// The command inputs bStop/bPark/bPower/bReset of FB_TelescopeControl (IAG50cm) are edge-triggered like the methods and are never
// written by the block; the block works on the request latches bStopActive/bParkActive/bPowerActive/bResetActive.
// Plan: BROTLib specs/plans/2026-11-09-iag50cm-command-model-unification.md, steps 1a/1b. One rig per test, one Scan() per PLC cycle.
FUNCTION_BLOCK IagCommandInputs_Tests EXTENDS TcUnit.FB_TestSuite
VAR
END_VAR

Held_Stop_Input_Stops_Once();
Park_Input_Edge_Parks_Like_Park();
Stop_Method_And_Input_Edge_In_One_Scan_Count_Once();
Power_Input_Is_Not_Written_By_The_Block();
Held_Slew_Input_Starts_The_Slew_Once();
Slew_Input_Falling_Does_Not_Abort_The_Slew();
Slew_Method_And_Input_Edge_In_One_Scan_Count_Once();
Slew_Input_In_The_Scan_Of_A_New_Error_Is_Rejected();
Track_Method_And_Track_Input_In_One_Scan_Count_Once();

// A held stop input is one command: one stop transaction, never repeated, never cleared by the block (IAG50cm command model step 1a).
METHOD PRIVATE Held_Stop_Input_Stops_Once
VAR_INST
	rig			: FB_IagRig;
	nStep		: INT;
	nCycles		: UINT;
	nEdges		: UINT;
	sTest		: STRING(80);
END_VAR
TEST('Held_Stop_Input_Stops_Once');
sTest := 'Held_Stop_Input_Stops_Once: ';
IF nStep >= 90 THEN
	RETURN;
END_IF
rig.Scan();
nCycles := nCycles + 1;
CASE nStep OF
0:	// wait for the clock, then power on
	IF rig.ClockValid THEN
		rig.fbTel.Init();
		nStep := 10;
		nCycles := 0;
	ELSIF nCycles > 2000 THEN
		AssertTrue(Condition := FALSE, Message := 'the astronomical clock never became valid');
		F_Note(bFailed := TRUE, sText := CONCAT(sTest, 'the astronomical clock never became valid'));
		nStep := 99;
		TEST_FINISHED();
	END_IF
10:	// wait until the startup has finished (READY_STATE 1.0)
	IF rig.Online THEN
		rig.fbTel.Slew(fAzimuth := 180.0, fAltitude := 45.0);
		nStep := 20;
		nCycles := 0;
	ELSIF nCycles > 1500 THEN
		AssertTrue(Condition := FALSE, Message := 'the mock telescope did not reach READY_STATE 1.0');
		F_Note(bFailed := TRUE, sText := CONCAT(sTest, 'the mock telescope did not reach READY_STATE 1.0'));
		nStep := 99;
		TEST_FINISHED();
	END_IF
20:	// an axis is moving
	IF rig.fbHa.MoveAxis OR rig.fbDec.MoveAxis THEN
		nCycles := 0;
		nStep := 30;
	ELSIF nCycles > 300 THEN
		AssertTrue(Condition := FALSE, Message := 'the slew did not start an axis move');
		F_Note(bFailed := TRUE, sText := CONCAT(sTest, 'the slew did not start an axis move'));
		nStep := 99;
		TEST_FINISHED();
	END_IF
30:	// a few scans of motion, then hold the stop INPUT (an ADS write, not the method)
	IF nCycles >= 5 THEN
		rig.SetStopInput(TRUE);
		nStep := 40;
		nCycles := 0;
	END_IF
40:	// the stop has settled: note the stop edges, keep holding the input
	IF NOT rig.fbTel.bStopActive AND rig.fbTel.bStopped AND nCycles > 5 THEN
		nEdges := rig.fbHa.nStopEdges + rig.fbDec.nStopEdges;
		AssertTrue(Condition := nEdges = 1, Message := 'the held input sent one stop to the moving axis');
		F_Note(bFailed := NOT (nEdges = 1), sText := CONCAT(sTest, 'the held input sent one stop to the moving axis'));
		nStep := 50;
		nCycles := 0;
	ELSIF nCycles > 400 THEN
		AssertTrue(Condition := FALSE, Message := 'the stop did not settle');
		F_Note(bFailed := TRUE, sText := CONCAT(sTest, 'the stop did not settle'));
		nStep := 99;
		TEST_FINISHED();
	END_IF
50:	// 60 more scans with the input still TRUE: no second stop, the latch stays down, the input is not cleared
	IF nCycles >= 60 THEN
		AssertTrue(Condition := rig.fbHa.nStopEdges + rig.fbDec.nStopEdges = nEdges, Message := 'a held input is not a second stop');
		F_Note(bFailed := NOT (rig.fbHa.nStopEdges + rig.fbDec.nStopEdges = nEdges), sText := CONCAT(sTest, 'a held input is not a second stop'));
		AssertTrue(Condition := NOT rig.fbTel.bStopActive, Message := 'the stop latch stayed down');
		F_Note(bFailed := NOT (NOT rig.fbTel.bStopActive), sText := CONCAT(sTest, 'the stop latch stayed down'));
		AssertTrue(Condition := rig.fbTel.bStop, Message := 'the block did not clear the input');
		F_Note(bFailed := NOT (rig.fbTel.bStop), sText := CONCAT(sTest, 'the block did not clear the input'));
		AssertTrue(Condition := rig.fbFocus.nStop = 1, Message := 'one stop for the focus');
		F_Note(bFailed := NOT (rig.fbFocus.nStop = 1), sText := CONCAT(sTest, 'one stop for the focus'));
		nStep := 99;
		TEST_FINISHED();
	END_IF
END_CASE
END_METHOD

// A rising park input starts the park exactly like Park(); the finished park is not replayed from the held input.
METHOD PRIVATE Park_Input_Edge_Parks_Like_Park
VAR_INST
	rig			: FB_IagRig;
	nStep		: INT;
	nCycles		: UINT;
	nEdges		: UINT;
	sTest		: STRING(80);
END_VAR
TEST('Park_Input_Edge_Parks_Like_Park');
sTest := 'Park_Input_Edge_Parks_Like_Park: ';
IF nStep >= 90 THEN
	RETURN;
END_IF
rig.Scan();
nCycles := nCycles + 1;
CASE nStep OF
0:	// wait for the clock, then power on
	IF rig.ClockValid THEN
		rig.fbTel.Init();
		nStep := 10;
		nCycles := 0;
	ELSIF nCycles > 2000 THEN
		AssertTrue(Condition := FALSE, Message := 'the astronomical clock never became valid');
		F_Note(bFailed := TRUE, sText := CONCAT(sTest, 'the astronomical clock never became valid'));
		nStep := 99;
		TEST_FINISHED();
	END_IF
10:	// wait until the startup has finished (READY_STATE 1.0)
	IF rig.Online THEN
		rig.SetParkInput(TRUE);
		nStep := 20;
		nCycles := 0;
	ELSIF nCycles > 1500 THEN
		AssertTrue(Condition := FALSE, Message := 'the mock telescope did not reach READY_STATE 1.0');
		F_Note(bFailed := TRUE, sText := CONCAT(sTest, 'the mock telescope did not reach READY_STATE 1.0'));
		nStep := 99;
		TEST_FINISHED();
	END_IF
20:	// the edge starts the park, as Park() would
	IF rig.fbTel.bParkActive THEN
		nStep := 30;
		nCycles := 0;
	ELSIF nCycles > 10 THEN
		AssertTrue(Condition := FALSE, Message := 'the park input edge did not start the park');
		F_Note(bFailed := TRUE, sText := CONCAT(sTest, 'the park input edge did not start the park'));
		nStep := 99;
		TEST_FINISHED();
	END_IF
30:
	IF rig.fbTel.bIsParked THEN
		nStep := 40;
		nCycles := 0;
	ELSIF nCycles > 3000 THEN
		AssertTrue(Condition := FALSE, Message := 'the park did not finish');
		F_Note(bFailed := TRUE, sText := CONCAT(sTest, 'the park did not finish'));
		nStep := 99;
		TEST_FINISHED();
	END_IF
40:	// the park ended with the input still TRUE: it is not replayed and not cleared
	IF nCycles >= 30 THEN
		AssertTrue(Condition := NOT rig.fbTel.bParkActive, Message := 'the park request ended');
		F_Note(bFailed := NOT (NOT rig.fbTel.bParkActive), sText := CONCAT(sTest, 'the park request ended'));
		AssertTrue(Condition := rig.fbTel.bIsParked, Message := 'the telescope stays parked');
		F_Note(bFailed := NOT (rig.fbTel.bIsParked), sText := CONCAT(sTest, 'the telescope stays parked'));
		AssertTrue(Condition := rig.fbTel.bPark, Message := 'the block did not clear the input');
		F_Note(bFailed := NOT (rig.fbTel.bPark), sText := CONCAT(sTest, 'the block did not clear the input'));
		nStep := 99;
		TEST_FINISHED();
	END_IF
END_CASE
END_METHOD

// Stop() and a stop input edge in one scan are one command (the method sets the edge memory).
METHOD PRIVATE Stop_Method_And_Input_Edge_In_One_Scan_Count_Once
VAR_INST
	rig			: FB_IagRig;
	nStep		: INT;
	nCycles		: UINT;
	nEdges		: UINT;
	sTest		: STRING(80);
END_VAR
TEST('Stop_Method_And_Input_Edge_In_One_Scan_Count_Once');
sTest := 'Stop_Method_And_Input_Edge_In_One_Scan_Count_Once: ';
IF nStep >= 90 THEN
	RETURN;
END_IF
rig.Scan();
nCycles := nCycles + 1;
CASE nStep OF
0:	// wait for the clock, then power on
	IF rig.ClockValid THEN
		rig.fbTel.Init();
		nStep := 10;
		nCycles := 0;
	ELSIF nCycles > 2000 THEN
		AssertTrue(Condition := FALSE, Message := 'the astronomical clock never became valid');
		F_Note(bFailed := TRUE, sText := CONCAT(sTest, 'the astronomical clock never became valid'));
		nStep := 99;
		TEST_FINISHED();
	END_IF
10:	// wait until the startup has finished (READY_STATE 1.0)
	IF rig.Online THEN
		rig.fbTel.Slew(fAzimuth := 180.0, fAltitude := 45.0);
		nStep := 20;
		nCycles := 0;
	ELSIF nCycles > 1500 THEN
		AssertTrue(Condition := FALSE, Message := 'the mock telescope did not reach READY_STATE 1.0');
		F_Note(bFailed := TRUE, sText := CONCAT(sTest, 'the mock telescope did not reach READY_STATE 1.0'));
		nStep := 99;
		TEST_FINISHED();
	END_IF
20:	// an axis is moving
	IF rig.fbHa.MoveAxis OR rig.fbDec.MoveAxis THEN
		nCycles := 0;
		nStep := 30;
	ELSIF nCycles > 300 THEN
		AssertTrue(Condition := FALSE, Message := 'the slew did not start an axis move');
		F_Note(bFailed := TRUE, sText := CONCAT(sTest, 'the slew did not start an axis move'));
		nStep := 99;
		TEST_FINISHED();
	END_IF
30:	// Stop() and the input edge in the same scan
	IF nCycles >= 5 THEN
		rig.fbTel.Stop();
		rig.SetStopInput(TRUE);
		nStep := 40;
		nCycles := 0;
	END_IF
40:
	IF NOT rig.fbTel.bStopActive AND rig.fbTel.bStopped AND nCycles > 5 THEN
		AssertTrue(Condition := rig.fbFocus.nStop = 1, Message := 'one Stop(): the focus stopped once');
		F_Note(bFailed := NOT (rig.fbFocus.nStop = 1), sText := CONCAT(sTest, 'one Stop(): the focus stopped once'));
		AssertTrue(Condition := rig.fbHa.nStopEdges + rig.fbDec.nStopEdges = 1, Message := 'one stop for the moving axis');
		F_Note(bFailed := NOT (rig.fbHa.nStopEdges + rig.fbDec.nStopEdges = 1), sText := CONCAT(sTest, 'one stop for the moving axis'));
		nStep := 99;
		TEST_FINISHED();
	ELSIF nCycles > 400 THEN
		AssertTrue(Condition := FALSE, Message := 'the stop did not settle');
		F_Note(bFailed := TRUE, sText := CONCAT(sTest, 'the stop did not settle'));
		nStep := 99;
		TEST_FINISHED();
	END_IF
END_CASE
END_METHOD

// A rising power input is an Init(); the block neither clears the input nor repeats the request.
METHOD PRIVATE Power_Input_Is_Not_Written_By_The_Block
VAR_INST
	rig			: FB_IagRig;
	nStep		: INT;
	nCycles		: UINT;
	nEdges		: UINT;
	sTest		: STRING(80);
END_VAR
TEST('Power_Input_Is_Not_Written_By_The_Block');
sTest := 'Power_Input_Is_Not_Written_By_The_Block: ';
IF nStep >= 90 THEN
	RETURN;
END_IF
rig.Scan();
nCycles := nCycles + 1;
CASE nStep OF
0:	// wait for the clock, then power on
	IF rig.ClockValid THEN
		rig.SetPowerInput(TRUE);
		nStep := 10;
		nCycles := 0;
	ELSIF nCycles > 2000 THEN
		AssertTrue(Condition := FALSE, Message := 'the astronomical clock never became valid');
		F_Note(bFailed := TRUE, sText := CONCAT(sTest, 'the astronomical clock never became valid'));
		nStep := 99;
		TEST_FINISHED();
	END_IF
10:	// wait until the startup has finished (READY_STATE 1.0)
	IF rig.Online THEN
		nStep := 20;
		nCycles := 0;
	ELSIF nCycles > 1500 THEN
		AssertTrue(Condition := FALSE, Message := 'the mock telescope did not reach READY_STATE 1.0');
		F_Note(bFailed := TRUE, sText := CONCAT(sTest, 'the mock telescope did not reach READY_STATE 1.0'));
		nStep := 99;
		TEST_FINISHED();
	END_IF
20:	// the power-on ran from the input edge and finished: the latch is down, the input is what the writer left
	IF nCycles >= 30 THEN
		AssertTrue(Condition := rig.Online, Message := 'the telescope is online');
		F_Note(bFailed := NOT (rig.Online), sText := CONCAT(sTest, 'the telescope is online'));
		AssertTrue(Condition := NOT rig.fbTel.bPowerActive, Message := 'the power-on request ended');
		F_Note(bFailed := NOT (NOT rig.fbTel.bPowerActive), sText := CONCAT(sTest, 'the power-on request ended'));
		AssertTrue(Condition := rig.fbTel.bPower, Message := 'the block did not clear the input');
		F_Note(bFailed := NOT (rig.fbTel.bPower), sText := CONCAT(sTest, 'the block did not clear the input'));
		nStep := 99;
		TEST_FINISHED();
	END_IF
END_CASE
END_METHOD

// A held slew input is one slew: it runs once and is neither repeated nor cleared by the block (command model step 1b).
METHOD PRIVATE Held_Slew_Input_Starts_The_Slew_Once
VAR_INST
	rig			: FB_IagRig;
	nStep		: INT;
	nCycles		: UINT;
	nEdges		: UINT;
	sTest		: STRING(80);
END_VAR
TEST('Held_Slew_Input_Starts_The_Slew_Once');
sTest := 'Held_Slew_Input_Starts_The_Slew_Once: ';
IF nStep >= 90 THEN
	RETURN;
END_IF
rig.Scan();
nCycles := nCycles + 1;
CASE nStep OF
0:	// wait for the clock, then power on
	IF rig.ClockValid THEN
		rig.fbTel.Init();
		nStep := 10;
		nCycles := 0;
	ELSIF nCycles > 2000 THEN
		AssertTrue(Condition := FALSE, Message := 'the astronomical clock never became valid');
		F_Note(bFailed := TRUE, sText := CONCAT(sTest, 'the astronomical clock never became valid'));
		nStep := 99;
		TEST_FINISHED();
	END_IF
10:	// wait until the startup has finished (READY_STATE 1.0)
	IF rig.Online THEN
		rig.SetSlewTargetInput(180.0, 45.0);
		rig.SetSlewInput(TRUE);
		nStep := 20;
		nCycles := 0;
	ELSIF nCycles > 1500 THEN
		AssertTrue(Condition := FALSE, Message := 'the mock telescope did not reach READY_STATE 1.0');
		F_Note(bFailed := TRUE, sText := CONCAT(sTest, 'the mock telescope did not reach READY_STATE 1.0'));
		nStep := 99;
		TEST_FINISHED();
	END_IF
20:	// an axis is moving
	IF rig.fbHa.MoveAxis OR rig.fbDec.MoveAxis THEN
		nCycles := 0;
		nStep := 30;
	ELSIF nCycles > 300 THEN
		AssertTrue(Condition := FALSE, Message := 'the slew did not start an axis move');
		F_Note(bFailed := TRUE, sText := CONCAT(sTest, 'the slew did not start an axis move'));
		nStep := 99;
		TEST_FINISHED();
	END_IF
30:	// the slew from the held input runs to its end
	IF NOT rig.fbTel.bSlewActive AND rig.fbTel.bStopped AND nCycles > 5 THEN
		nStep := 40;
		nCycles := 0;
	ELSIF nCycles > 3000 THEN
		AssertTrue(Condition := FALSE, Message := 'the slew did not finish');
		F_Note(bFailed := TRUE, sText := CONCAT(sTest, 'the slew did not finish'));
		nStep := 99;
		TEST_FINISHED();
	END_IF
40:	// 60 scans with the input still TRUE: the slew is not started again, the input is not cleared
	IF nCycles >= 60 THEN
		AssertTrue(Condition := NOT rig.fbTel.bSlewActive, Message := 'the slew was not restarted');
		F_Note(bFailed := NOT (NOT rig.fbTel.bSlewActive), sText := CONCAT(sTest, 'the slew was not restarted'));
		AssertTrue(Condition := rig.fbTel.TCS_command <> E_TCSCommand.slew, Message := 'no slew command is running');
		F_Note(bFailed := NOT (rig.fbTel.TCS_command <> E_TCSCommand.slew), sText := CONCAT(sTest, 'no slew command is running'));
		AssertTrue(Condition := rig.fbTel.bSlew, Message := 'the block did not clear the input');
		F_Note(bFailed := NOT (rig.fbTel.bSlew), sText := CONCAT(sTest, 'the block did not clear the input'));
		nStep := 99;
		TEST_FINISHED();
	END_IF
END_CASE
END_METHOD

// The slew input falling does not abort the slew; it ends only by its own completion or a stop.
METHOD PRIVATE Slew_Input_Falling_Does_Not_Abort_The_Slew
VAR_INST
	rig			: FB_IagRig;
	nStep		: INT;
	nCycles		: UINT;
	nEdges		: UINT;
	sTest		: STRING(80);
END_VAR
TEST('Slew_Input_Falling_Does_Not_Abort_The_Slew');
sTest := 'Slew_Input_Falling_Does_Not_Abort_The_Slew: ';
IF nStep >= 90 THEN
	RETURN;
END_IF
rig.Scan();
nCycles := nCycles + 1;
CASE nStep OF
0:	// wait for the clock, then power on
	IF rig.ClockValid THEN
		rig.fbTel.Init();
		nStep := 10;
		nCycles := 0;
	ELSIF nCycles > 2000 THEN
		AssertTrue(Condition := FALSE, Message := 'the astronomical clock never became valid');
		F_Note(bFailed := TRUE, sText := CONCAT(sTest, 'the astronomical clock never became valid'));
		nStep := 99;
		TEST_FINISHED();
	END_IF
10:	// wait until the startup has finished (READY_STATE 1.0)
	IF rig.Online THEN
		rig.SetSlewTargetInput(180.0, 45.0);
		rig.SetSlewInput(TRUE);
		nStep := 20;
		nCycles := 0;
	ELSIF nCycles > 1500 THEN
		AssertTrue(Condition := FALSE, Message := 'the mock telescope did not reach READY_STATE 1.0');
		F_Note(bFailed := TRUE, sText := CONCAT(sTest, 'the mock telescope did not reach READY_STATE 1.0'));
		nStep := 99;
		TEST_FINISHED();
	END_IF
20:	// an axis is moving
	IF rig.fbHa.MoveAxis OR rig.fbDec.MoveAxis THEN
		nCycles := 0;
		nStep := 25;
	ELSIF nCycles > 300 THEN
		AssertTrue(Condition := FALSE, Message := 'the slew did not start an axis move');
		F_Note(bFailed := TRUE, sText := CONCAT(sTest, 'the slew did not start an axis move'));
		nStep := 99;
		TEST_FINISHED();
	END_IF
25:	// the writer drops the input while the axis moves
	IF nCycles >= 5 THEN
		rig.SetSlewInput(FALSE);
		nStep := 30;
		nCycles := 0;
	END_IF
30:
	IF nCycles >= 5 THEN
		AssertTrue(Condition := rig.fbTel.bSlewActive, Message := 'the slew goes on after the input fell');
		F_Note(bFailed := NOT (rig.fbTel.bSlewActive), sText := CONCAT(sTest, 'the slew goes on after the input fell'));
		nStep := 40;
		nCycles := 0;
	END_IF
40:
	IF NOT rig.fbTel.bSlewActive AND rig.fbTel.bStopped AND nCycles > 5 THEN
		nStep := 99;
		TEST_FINISHED();
	ELSIF nCycles > 3000 THEN
		AssertTrue(Condition := FALSE, Message := 'the slew did not finish');
		F_Note(bFailed := TRUE, sText := CONCAT(sTest, 'the slew did not finish'));
		nStep := 99;
		TEST_FINISHED();
	END_IF
END_CASE
END_METHOD

// Slew() and a slew input edge in one scan are one slew (the method sets the edge memory).
METHOD PRIVATE Slew_Method_And_Input_Edge_In_One_Scan_Count_Once
VAR_INST
	rig			: FB_IagRig;
	nStep		: INT;
	nCycles		: UINT;
	nEdges		: UINT;
	sTest		: STRING(80);
END_VAR
TEST('Slew_Method_And_Input_Edge_In_One_Scan_Count_Once');
sTest := 'Slew_Method_And_Input_Edge_In_One_Scan_Count_Once: ';
IF nStep >= 90 THEN
	RETURN;
END_IF
rig.Scan();
nCycles := nCycles + 1;
CASE nStep OF
0:	// wait for the clock, then power on
	IF rig.ClockValid THEN
		rig.fbTel.Init();
		nStep := 10;
		nCycles := 0;
	ELSIF nCycles > 2000 THEN
		AssertTrue(Condition := FALSE, Message := 'the astronomical clock never became valid');
		F_Note(bFailed := TRUE, sText := CONCAT(sTest, 'the astronomical clock never became valid'));
		nStep := 99;
		TEST_FINISHED();
	END_IF
10:	// wait until the startup has finished (READY_STATE 1.0)
	IF rig.Online THEN
		rig.fbTel.Slew(fAzimuth := 180.0, fAltitude := 45.0);
		rig.SetSlewInput(TRUE);
		nStep := 20;
		nCycles := 0;
	ELSIF nCycles > 1500 THEN
		AssertTrue(Condition := FALSE, Message := 'the mock telescope did not reach READY_STATE 1.0');
		F_Note(bFailed := TRUE, sText := CONCAT(sTest, 'the mock telescope did not reach READY_STATE 1.0'));
		nStep := 99;
		TEST_FINISHED();
	END_IF
20:	// an axis is moving
	IF rig.fbHa.MoveAxis OR rig.fbDec.MoveAxis THEN
		nCycles := 0;
		nStep := 30;
	ELSIF nCycles > 300 THEN
		AssertTrue(Condition := FALSE, Message := 'the slew did not start an axis move');
		F_Note(bFailed := TRUE, sText := CONCAT(sTest, 'the slew did not start an axis move'));
		nStep := 99;
		TEST_FINISHED();
	END_IF
30:
	IF NOT rig.fbTel.bSlewActive AND rig.fbTel.bStopped AND nCycles > 5 THEN
		nStep := 40;
		nCycles := 0;
	ELSIF nCycles > 3000 THEN
		AssertTrue(Condition := FALSE, Message := 'the slew did not finish');
		F_Note(bFailed := TRUE, sText := CONCAT(sTest, 'the slew did not finish'));
		nStep := 99;
		TEST_FINISHED();
	END_IF
40:	IF nCycles >= 60 THEN
		AssertTrue(Condition := NOT rig.fbTel.bSlewActive, Message := 'no second slew');
		F_Note(bFailed := NOT (NOT rig.fbTel.bSlewActive), sText := CONCAT(sTest, 'no second slew'));
		AssertTrue(Condition := rig.fbHa.nStopEdges + rig.fbDec.nStopEdges = 0, Message := 'no restart stop');
		F_Note(bFailed := NOT (rig.fbHa.nStopEdges + rig.fbDec.nStopEdges = 0), sText := CONCAT(sTest, 'no restart stop'));
		nStep := 99;
		TEST_FINISHED();
	END_IF
END_CASE
END_METHOD

// D1 (template body step S1.d): a slew input edge in the scan of a new axis error is rejected at arrival (the gate sees this scan's error), not accepted and dropped silently.
METHOD PRIVATE Slew_Input_In_The_Scan_Of_A_New_Error_Is_Rejected
VAR_INST
	rig			: FB_IagRig;
	nStep		: INT;
	nCycles		: UINT;
	sTest		: STRING(80);
END_VAR
TEST('Slew_Input_In_The_Scan_Of_A_New_Error_Is_Rejected');
sTest := 'Slew_Input_In_The_Scan_Of_A_New_Error_Is_Rejected: ';
IF nStep >= 90 THEN
	RETURN;
END_IF
rig.Scan();
nCycles := nCycles + 1;
CASE nStep OF
0:	// wait for the clock, then power on
	IF rig.ClockValid THEN
		rig.fbTel.Init();
		nStep := 10;
		nCycles := 0;
	ELSIF nCycles > 2000 THEN
		AssertTrue(Condition := FALSE, Message := 'the astronomical clock never became valid');
		F_Note(bFailed := TRUE, sText := CONCAT(sTest, 'the astronomical clock never became valid'));
		nStep := 99;
		TEST_FINISHED();
	END_IF
10:	// wait until the startup has finished (READY_STATE 1.0)
	IF rig.Online THEN
		rig.SetHorizon(-90.0);
		rig.SetSafeAltitude(-90.0);
		rig.SetSlewTargetInput(fAzimuth := 180.0, fAltitude := 45.0);
		rig.InjectHaError(16#4550);
		rig.SetSlewInput(TRUE);
		nStep := 20;
		nCycles := 0;
	ELSIF nCycles > 1500 THEN
		AssertTrue(Condition := FALSE, Message := 'the mock telescope did not reach READY_STATE 1.0');
		F_Note(bFailed := TRUE, sText := CONCAT(sTest, 'the mock telescope did not reach READY_STATE 1.0'));
		nStep := 99;
		TEST_FINISHED();
	END_IF
20:	// the slew edge came in the scan in which the axis error appeared: rejected at arrival, with a log, nothing latched
	IF nCycles >= 5 THEN
		AssertTrue(Condition := rig.fbTel.bError, Message := 'the error is reported');
		F_Note(bFailed := NOT (rig.fbTel.bError), sText := CONCAT(sTest, 'the error is reported'));
		AssertTrue(Condition := rig.fbTel.nCommandRejectCount >= 1, Message := 'the slew was rejected and counted');
		F_Note(bFailed := NOT (rig.fbTel.nCommandRejectCount >= 1), sText := CONCAT(sTest, 'the slew was rejected and counted'));
		AssertTrue(Condition := NOT rig.fbTel.bSlewActive, Message := 'no slew is latched');
		F_Note(bFailed := NOT (NOT rig.fbTel.bSlewActive), sText := CONCAT(sTest, 'no slew is latched'));
		nStep := 99;
		TEST_FINISHED();
	END_IF
END_CASE
END_METHOD

// D4 (template body step S1.f): Track() and a bTrack input edge in one scan are one command (Track() marks the edge memory of the track input), as in MONETcommon.
METHOD PRIVATE Track_Method_And_Track_Input_In_One_Scan_Count_Once
VAR_INST
	rig			: FB_IagRig;
	nStep		: INT;
	nCycles		: UINT;
	sTest		: STRING(80);
END_VAR
TEST('Track_Method_And_Track_Input_In_One_Scan_Count_Once');
sTest := 'Track_Method_And_Track_Input_In_One_Scan_Count_Once: ';
IF nStep >= 90 THEN
	RETURN;
END_IF
rig.Scan();
nCycles := nCycles + 1;
CASE nStep OF
0:	// wait for the clock, then power on
	IF rig.ClockValid THEN
		rig.fbTel.Init();
		nStep := 10;
		nCycles := 0;
	ELSIF nCycles > 2000 THEN
		AssertTrue(Condition := FALSE, Message := 'the astronomical clock never became valid');
		F_Note(bFailed := TRUE, sText := CONCAT(sTest, 'the astronomical clock never became valid'));
		nStep := 99;
		TEST_FINISHED();
	END_IF
10:	// wait until the startup has finished (READY_STATE 1.0)
	IF rig.Online THEN
		rig.SetHorizon(-90.0);
		rig.SetSafeAltitude(-90.0);
		rig.fbTel.Track(fRightAscension := 100.0, fDeclination := 30.0);
		rig.SetTrackInput(TRUE);
		nStep := 20;
		nCycles := 0;
	ELSIF nCycles > 1500 THEN
		AssertTrue(Condition := FALSE, Message := 'the mock telescope did not reach READY_STATE 1.0');
		F_Note(bFailed := TRUE, sText := CONCAT(sTest, 'the mock telescope did not reach READY_STATE 1.0'));
		nStep := 99;
		TEST_FINISHED();
	END_IF
20:	// one command: the goto of Track() runs, the bTrack edge of the same scan is not a second (replacing) command
	IF nCycles = 3 THEN
		AssertTrue(Condition := rig.fbTel.bGotoActive, Message := 'the goto of Track() is latched');
		F_Note(bFailed := NOT (rig.fbTel.bGotoActive), sText := CONCAT(sTest, 'the goto of Track() is latched'));
		AssertTrue(Condition := NOT rig.fbTel.bTrackActive, Message := 'the input edge did not replace it');
		F_Note(bFailed := NOT (NOT rig.fbTel.bTrackActive), sText := CONCAT(sTest, 'the input edge did not replace it'));
		AssertTrue(Condition := rig.fbTel.nCommandRejectCount = 0, Message := 'nothing was rejected');
		F_Note(bFailed := NOT (rig.fbTel.nCommandRejectCount = 0), sText := CONCAT(sTest, 'nothing was rejected'));
		AssertTrue(Condition := NOT rig.fbTel.bMoveAbortPending, Message := 'no abort stop for a replacement');
		F_Note(bFailed := NOT (NOT rig.fbTel.bMoveAbortPending), sText := CONCAT(sTest, 'no abort stop for a replacement'));
		nStep := 99;
		TEST_FINISHED();
	END_IF
END_CASE
END_METHOD

END_FUNCTION_BLOCK

(* stored: Version 1.1.0.1, ProductVersion 3.1.4024.15
   POU IagCommandInputs_Tests: Id {ce2b8202-2582-4506-8c21-3f082b0ac712}, SpecialFunc None
   Method Held_Stop_Input_Stops_Once: Id {e863a4e4-6e59-4764-bafa-ca5df7d13b80}
   Method Park_Input_Edge_Parks_Like_Park: Id {f17494b3-cf10-46c0-8483-234010719e5d}
   Method Stop_Method_And_Input_Edge_In_One_Scan_Count_Once: Id {29a08ce9-a108-4305-b65a-c0856bef6315}
   Method Power_Input_Is_Not_Written_By_The_Block: Id {fe2277a3-6300-45d2-a7e1-b017000bfbfe}
   Method Held_Slew_Input_Starts_The_Slew_Once: Id {131a17aa-45da-4c24-9ff5-93bdb4077968}
   Method Slew_Input_Falling_Does_Not_Abort_The_Slew: Id {b71c0bc3-66bd-4cd1-bea4-eebc87eab3d2}
   Method Slew_Method_And_Input_Edge_In_One_Scan_Count_Once: Id {4ef17647-4434-4785-ab0d-f642668748f4}
   Method Slew_Input_In_The_Scan_Of_A_New_Error_Is_Rejected: Id {8dd2e7da-81e6-46be-a6f4-4090ce41f783}
   Method Track_Method_And_Track_Input_In_One_Scan_Count_Once: Id {de0f8ee8-46f6-484c-b809-bda86120714e} *)
